(* IEC 61131-3 sources: SortJet_MasterSPS_Aufbau.fbsproj/09_Station/UnterStationsbausteine, 8 files *)

(* ---- Geblaese_Schuetz_FB_V01_00_00.fb.st ---- *)
(* METADATA
{
	"v3Meta": {
		"objectGuid": "c9895c16-daf8-42f8-8f64-ac96a02bd793"
	}
}
*)
FUNCTION_BLOCK Geblaese_Schuetz_FB_V01_00_00
VAR_INPUT

  // BOOLEAN
  bpAktivieren              : BOOL;
  bpStart                   : BOOL;
  bpReset                   : BOOL;
  bpFreigabe                : BOOL;
  bpTeilnehmerErreichbar    : BOOL := TRUE;
  bpIOsBoschDrive               : BOOL;

  // EINGÄNGE
  bpMotorschutzschalter_OK  : BOOL;
  bpDrehzahlErreicht        : BOOL := TRUE; // Sanftanlauf: Drehzahl erreicht (ohne Sanftanlauf TRUE lassen)

  // DROSSELKLAPPE
  bpDrosselklappeAnforderung : BOOL; // Station: Drosselklappe soll offen sein (Transport, Anlegen, Geblaese gestartet)

  // STEUERUNG (wann das Geblaese laufen soll, Aktion Steuerung)
  bpAutomatik        : BOOL;            // Automatik / Check: Geblaese nach Aktivitaet mit Energiesparmodus
  bpAktivitaet       : BOOL;            // Station braucht das Geblaese (z.B. Auftrag aktiv)
  bpAktivitaetFlanke : BOOL;            // Anlegestation: nur die steigende Flanke der Aktivitaet startet, danach Abschaltzeit
  bpTaster           : BOOL;            // Taster am Geblaese: umschalten
  bpHandEin          : BOOL;            // Handbetrieb: Geblaese laeuft, solange gesetzt
  bpSperre           : BOOL;            // Geblaese sofort aus (Reset, Verriegelung)
  tpMindestlaufzeit  : TIME := T#500MS; // Der Taster schaltet erst nach dieser Laufzeit aus

  // STRUKT
  stStationsNummern       : Station_ST;

END_VAR
VAR_OUTPUT

  // BOOLEAN
  bpFehler                 : BOOL;
  bpDone                   : BOOL;
  bpStarteGeblaese         : BOOL; // Geblaese wird angesteuert (Schuetz)
  bpDrosselklappeOeffnen   : BOOL; // Drosselklappe oeffnen: angefordert und Geblaese laeuft

  // WORD
  wpFehlerNr : Fehlerkonstanten_EN;

END_VAR
VAR

  // BOOLEAN
  blErsterZyklus           : BOOL := TRUE; // Initialisierung
  blMeldungAbgesetzt       : BOOL := FALSE;
  blMotorschutzschalter_OK : BOOL;

  // ARRAY
  awlErrorAdditional : ARRAY [0..25]  OF WORD;

  // STEPS
  steplStart      : Steps_TE;

  // TIMER
  tonlStartGeblaese          : TON;
  tonlWarteAufGeblaeseLaeuft : TON;
  toflWarteAufWiederAnlauf   : TOF;
  toflMotorschutz            : TOF;
  toflEnergiesparModus       : TOF; // Energiesparmodus: Geblaese nach der Abschaltzeit ohne Aktivitaet aus
  tonlMindestlaufzeit        : TON;

  // TRIGGER
  rtlAutomatik               : R_TRIG;
  rtlAktivitaet              : R_TRIG;
  rtlTaster                  : R_TRIG;

  // BOOLEAN (Steuerung)
  blTasterAus                : BOOL; // Automatik: Geblaese per Taster ausgeschaltet (bis zur naechsten Aktivitaet)
  blHandTaster               : BOOL; // Handbetrieb: Geblaese per Taster eingeschaltet

END_VAR
VAR

  // HARDWARE EINGAENGE
  in_bMotorschutzschalter_OK    AT %I* : BOOL;

  // HARDWARE AUSGAENGE
  out_bStarteGeblaese           AT %Q* : BOOL;

END_VAR

VAR CONSTANT

  // TIME
  WARTEZEIT_BIS_WIEDERANLAUF          : TIME := T#7000MS;
  WARTEZEIT_BIS_GEBLAESE_HOCHGELAUFEN : TIME := T#2000MS;

END_VAR

//-------------------------------------------------------------------------------------------------
// BAUSTEIN: INITIALISIERUNG
//-------------------------------------------------------------------------------------------------
IF ( blErsterZyklus ) THEN
  blErsterZyklus:=FALSE;

  (* Hinweis:
     - Timer initialisieren
  *)
  toflWarteAufWiederAnlauf(IN:=FALSE);
  tonlWarteAufGeblaeseLaeuft(IN:=FALSE);

END_IF
// IO Zuweisung
IF ( bpIOsBoschDrive ) THEN
  blMotorschutzschalter_OK  := bpMotorschutzschalter_OK;
ELSE
  blMotorschutzschalter_OK  := in_bMotorschutzschalter_OK;
END_IF

//-------------------------------------------------------------------------------------------------
// BAUSTEIN: DEAKTIVIEREN
//-------------------------------------------------------------------------------------------------
IF ( NOT bpAktivieren ) THEN
  bpDone                 := TRUE;
  bpStarteGeblaese       := FALSE;
  bpDrosselklappeOeffnen := FALSE;
  bpFehler   := FALSE;
  wpFehlerNr := cMELDUNG_NULL;

  RETURN;

END_IF

//-------------------------------------------------------------------------------------------------
// BAUSTEIN: STEUERUNG
//-------------------------------------------------------------------------------------------------
Steuerung();

//-------------------------------------------------------------------------------------------------
// BAUSTEIN: TIMER
//-------------------------------------------------------------------------------------------------
toflWarteAufWiederAnlauf(IN :=     out_bStarteGeblaese,
                          PT := WARTEZEIT_BIS_WIEDERANLAUF);

tonlWarteAufGeblaeseLaeuft(IN :=     out_bStarteGeblaese,
                            PT := WARTEZEIT_BIS_GEBLAESE_HOCHGELAUFEN );

toflMotorschutz( IN := blMotorschutzschalter_OK, PT := T#5S );

(* Hinweis:
   - Einschaltverzoegerung
*)
tonlStartGeblaese(IN :=     bpStart
                   AND bpFreigabe
                   AND NOT toflWarteAufWiederAnlauf.Q
                   AND NOT bpReset,
                   PT := T#0S);

//-------------------------------------------------------------------------------------------------
// BAUSTEIN: STEUERUNG
//-------------------------------------------------------------------------------------------------
IF ( bpReset ) THEN

  bpStart   := FALSE;
  bpDone    := FALSE;
  bpReset   := FALSE;
  bpFehler  := FALSE;

  blMeldungAbgesetzt := FALSE;

  wpFehlerNr := cMELDUNG_NULL;

  out_bStarteGeblaese := FALSE;

ELSE
  Start();
  Meldungen();

END_IF

//-------------------------------------------------------------------------------------------------
// BAUSTEIN: AUSGAENGE
//-------------------------------------------------------------------------------------------------
(* Hinweis:
   - Ansteuerung des Geblaeses fuer Stationen, die den Ausgang selbst schalten (z.B. zwei Geblaese oder Ausgang am Umrichter)
   - Die Drosselklappe ist nur offen, wenn sie angefordert ist und das Geblaese laeuft (Drehzahl erreicht)
*)
bpStarteGeblaese       := out_bStarteGeblaese;
bpDrosselklappeOeffnen := bpDrosselklappeAnforderung AND bpDone;
END_FUNCTION_BLOCK

(* ---- Hub_FB_V01_00_00.fb.st ---- *)
(* METADATA
{
	"v3Meta": {
		"objectGuid": "03cf6ff6-d378-4ff5-8445-541e648ef0b8"
	}
}
*)
FUNCTION_BLOCK Hub_FB_V01_00_00
VAR_INPUT

  // BOOLEAN
  bpAktivieren               : BOOL;
  bpStartHubAuf              : BOOL;
  bpStartHubAb               : BOOL;
  bpReset                    : BOOL;
  bpSensorEinlaufNachfolger  : BOOL;
  bpSensorAuslaufVorgaenger  : BOOL;
  bpSensorEinlauf            : BOOL;
  bpSensorAuslauf            : BOOL;

  // STRUCT
  stStationsNummern          : Station_ST;

END_VAR
VAR_OUTPUT

  // BOOLEAN
  bpFehler        : BOOL;
  bpDone          : BOOL;

  // WORD
  wpFehlerNr : Fehlerkonstanten_EN;

  // ENUM
  epHubStatus  : Hub_EN; // Status: Gibt die Aktuelle Position des Antriebs aus

END_VAR

VAR

  // BOOLEAN
  blErsterZyklus        : BOOL := TRUE;

  // TIMER
  tonlMaxWarteZeit                        : TON;
  tonlHubAntriebOK                        : TON;
  tonlMaximaleWartezeitAufReset           : TON;
  tonlFehlermeldungUnterdrueckenAntriebOK : TON;
  tonlReset                               : TON;

  // STEPS
  steplHubAb    : Steps_TE;
  steplHubAuf   : Steps_TE;
  steplReset    : Steps_TE;

END_VAR

VAR
  // HARDWARE EINGÄNGE
  in_bSensorNichtUnten             AT%I* : BOOL;
  in_bSensorNichtOben              AT%I* : BOOL;
  in_bMotorstarter_OK              AT%I* : BOOL;
  in_bLSBremse_OK                  AT%I* : BOOL;
  in_bLS400V_OK                    AT%I* : BOOL;

  // HARDWARE AUSGÄNGE
  out_bHubAbSetzen                 AT%Q* : BOOL;
  out_bHubAufSetzen                AT%Q* : BOOL;
  out_bReset                       AT%Q* : BOOL;
  out_bBremseLoesen                AT%Q* : BOOL;

END_VAR

VAR CONSTANT

  // TIME
  MAXIMALE_WARTEZEIT_HUB                       : TIME := T#5000MS; // Maximale Wartezeit die abgewartet wird bis der Hub-Antrieb auf Position gefahren ist

END_VAR
//-------------------------------------------------------------------------------------------------
// BAUSTEIN: INITIALISIERUNG
//-------------------------------------------------------------------------------------------------
IF ( blErsterZyklus ) THEN
  blErsterZyklus := FALSE;

  (* Hinweis:
     - Timer initialisieren
  *)
  tonlHubAntriebOK(IN:=TRUE);
  tonlMaxWarteZeit(IN:=FALSE);
  tonlFehlermeldungUnterdrueckenAntriebOK( IN := FALSE );

END_IF

//-------------------------------------------------------------------------------------------------
// BAUSTEIN: AKTIONEN
//-------------------------------------------------------------------------------------------------
IF ( bpAktivieren ) THEN

  HubAuf();
  HubAb();

  Ausgaenge();
  Meldungen();
  Timer();
  Reset();

ELSE

  bpDone   := TRUE;
  bpFehler := FALSE;

  IF (bpStartHubAb AND NOT bpStartHubAuf) THEN
    epHubStatus := eHub_Unten;
  ELSIF (bpStartHubAuf AND NOT bpStartHubAb) THEN
    epHubStatus := eHub_Oben;
  ELSIF (bpStartHubAb AND NOT bpStartHubAuf) THEN
    epHubStatus := eHub_Undefiniert;
  END_IF

END_IF
END_FUNCTION_BLOCK

(* ---- Transportsperre_Foerderbaender_FB_V01_00_00.fb.st ---- *)
(* METADATA
{
	"v3Meta": {
		"objectGuid": "85c14a01-ee4c-4a24-bcca-8fef195064c0"
	}
}
*)
{attribute 'excludefrombuild'}
FUNCTION_BLOCK Transportsperre_Foerderbaender_FB_V01_00_00
VAR_INPUT

  // HARDWARE EINGAENGE
  in_bOben            : BOOL; // STATUS: Sensor meldt ausgfahren  [Oben]

  // BOOLEAN
  bpAktivieren        : BOOL;
  bpStartRunter       : BOOL; // BETRIEBTYP: Zylinder wird ausgefahren
  bpStartHoch         : BOOL; // BETRIEBTYP: Zylinder wird eingefahren
  bpReset             : BOOL; // BETRIEBTYP: Zylinderbaustein wird zurueckgesetzt
  bpFreigabe          : BOOL;

  // OPTIONEN
  bpAbfrageObenVorhanden  : BOOL := TRUE;   // Endlagensensor oben vorhanden, sonst gilt die Endlage nach tpBewegungszeit
  bpAbfrageUntenVorhanden : BOOL := TRUE;   // Endlagensensor unten vorhanden, sonst gilt die Endlage nach tpBewegungszeit
  tpBewegungszeit         : TIME := T#800MS; // Bewegungszeit je Richtung ohne Endlagensensor

END_VAR
VAR_OUTPUT

  // BOOLEAN
  bpFehler            : BOOL;
  bpDone              : BOOL;

  // WORD
  wpFehlerNr          : Fehlerkonstanten_EN;

  // ENUM
  wpStatus            : TransportsperrenStatus_EN;

END_VAR
VAR
  // STEPS
  steplHoch         : Steps_TE;
  steplRunter       : Steps_TE;

  // TIMER
  tonlOben                 : TON; // EINSCHALTVERZOEGERUNG: Warten bis der Zylinder eingefahren wurde. Sonst wird ein Fehlerausgegeben
  tonlUnten                : TON; // EINSCHALTVERZOEGERUNG: Warten bis der Zylinder ausgefahren wurde. Sonst wird ein Fehlerausgegeben
  tonlBewegungszeitHoch    : TON; // Bewegungszeit ohne Endlagensensor oben
  tonlBewegungszeitRunter  : TON; // Bewegungszeit ohne Endlagensensor unten
  tofHoch                  : TOF;
  tofRunter                : TOF;

END_VAR

VAR

  // HARDWARE EINGAENGE
  in_bUnten     AT %I* : BOOL; // STATUS: Sensor meldt eingefahren [Unten]

  // HARDWARE AUSGAENGE
  out_bRunter   AT %Q* : BOOL; // AKTION: Zylinder einfahren

END_VAR
VAR CONSTANT

  // TIME
  cZEITLICHE_UEBERWACHUNG_BEWEGUNG_ZYLINDER : TIME := T#15s;

END_VAR
(* Hinweis:
   - Ein Ausgang (Federrueckstell- Ventil): Runter haelt den Ausgang, Hoch nimmt ihn zurueck
*)

//-------------------------------------------------------------------------------------------------
// BAUSTEIN: RESET / DEAKTIVIERT
//-------------------------------------------------------------------------------------------------
(* Hinweis:
   - Reset oder deaktiviert: Ausgang aus, Ketten und Timer zuruecksetzen, Done und Fehler loeschen
   - Der Baustein setzt bpReset selbst zurueck, der Aufrufer wartet nicht auf Done
   - Ein deaktivierter Baustein meldet kein Done; der Aufrufer verknuepft das Warten auf Done
     mit der Aktivierung aus der MK (z.B. Transportsperre.bpDone OR NOT stStationsAufbau.bX)
*)
IF ( bpReset OR NOT bpAktivieren ) THEN

  out_bRunter := FALSE;

  bpStartRunter := FALSE;
  bpStartHoch   := FALSE;

  steplHoch   := STEP_0_E;
  steplRunter := STEP_0_E;

  tonlOben( IN := FALSE );
  tonlUnten( IN := FALSE );
  tonlBewegungszeitHoch( IN := FALSE );
  tonlBewegungszeitRunter( IN := FALSE );
  tofHoch( IN := FALSE );
  tofRunter( IN := FALSE );

  bpDone     := FALSE;
  bpFehler   := FALSE;
  wpFehlerNr := cMELDUNG_NULL;

  bpReset := FALSE;

  RETURN;

END_IF

//-------------------------------------------------------------------------------------------------
// BAUSTEIN: AKTIONEN
//-------------------------------------------------------------------------------------------------
HochFahren();
RunterFahren();

// Umschaltpause zwischen den Richtungen
tofHoch( IN := bpStartHoch, PT := T#1S );
tofRunter( IN := bpStartRunter, PT := T#1S );

//-------------------------------------------------------------------------------------------------
// STATUS DER TRANSPORTSPERRE
//-------------------------------------------------------------------------------------------------
(* Hinweis:
   - Status aus der Sensorik, soweit Endlagensensoren vorhanden sind
   - Ohne Sensor bleibt der Status, den die Schrittketten nach der Bewegungszeit setzen
*)
IF ( bpAbfrageObenVorhanden AND bpAbfrageUntenVorhanden ) THEN

  IF (     in_bOben
       AND NOT in_bUnten )
  THEN
    wpStatus := eTransportsperreOben;
  ELSIF(   in_bUnten
         AND NOT in_bOben )
  THEN
    wpStatus := eTransportsperreUnten;
  ELSE
    wpStatus := eTransportsperreUndefiniert;
  END_IF

ELSIF ( bpAbfrageObenVorhanden ) THEN

  IF ( in_bOben ) THEN
    wpStatus := eTransportsperreOben;
  ELSIF ( wpStatus = eTransportsperreOben ) THEN
    wpStatus := eTransportsperreUndefiniert;
  END_IF

ELSIF ( bpAbfrageUntenVorhanden ) THEN

  IF ( in_bUnten ) THEN
    wpStatus := eTransportsperreUnten;
  ELSIF ( wpStatus = eTransportsperreUnten ) THEN
    wpStatus := eTransportsperreUndefiniert;
  END_IF

END_IF
END_FUNCTION_BLOCK

(* ---- Transportsperre_Kipptisch_FB_V01_00_00.fb.st ---- *)
(* METADATA
{
	"v3Meta": {
		"objectGuid": "32d63b77-62b3-4c1f-9a6d-0b9e7860b01c"
	}
}
*)
{attribute 'excludefrombuild'}
FUNCTION_BLOCK Transportsperre_Kipptisch_FB_V01_00_00
VAR_INPUT

  // BOOLEAN
  bpAktivieren        : BOOL;
  bpStartAusfahren    : BOOL; // BETRIEBTYP: Zylinder wird ausgefahren
  bpStartEinfahren    : BOOL; // BETRIEBTYP: Zylinder wird eingefahren
  bpReset             : BOOL; // BETRIEBTYP: Zylinderbaustein wird zurueckgesetzt
  bpFreigabe          : BOOL; //
  bpFreigabeEinfahren : BOOL; // Freigabe von der Folgestation, dass die Sperre runter fahren darf

  // OPTIONEN
  bpAbfrageAusgefahrenVorhanden : BOOL := TRUE;   // Endlagensensor ausgefahren vorhanden, sonst gilt die Endlage nach tpBewegungszeit
  bpAbfrageEingefahrenVorhanden : BOOL := TRUE;   // Endlagensensor eingefahren vorhanden, sonst gilt die Endlage nach tpBewegungszeit
  tpBewegungszeit               : TIME := T#800MS; // Bewegungszeit je Richtung ohne Endlagensensor

END_VAR
VAR_OUTPUT

  // BOOLEAN
  bpFehler            : BOOL;
  bpDone              : BOOL;
  bpFreigabeKippen    : BOOL;
  bpFreigabeTransport : BOOL;

  // WORD
  wpFehlerNr       : Fehlerkonstanten_EN;

  // ENUM
  wpStatusZylinder : PneumatikZylinderStatus_EN;

END_VAR
VAR
  // STEPS
  steplAusfahren   : Steps_TE;
  steplEinfahren   : Steps_TE;

  // TIMER
  tonlZylinderEingefahren    : TON; // EINSCHALTVERZOEGERUNG: Warten bis der Zylinder eingefahren wurde. Sonst wird ein Fehlerausgegeben
  tonlZylinderAusgefahren    : TON; // EINSCHALTVERZOEGERUNG: Warten bis der Zylinder ausgefahren wurde. Sonst wird ein Fehlerausgegeben
  tonlBewegungszeitEinfahren : TON; // Bewegungszeit ohne Endlagensensor eingefahren
  tonlBewegungszeitAusfahren : TON; // Bewegungszeit ohne Endlagensensor ausgefahren
  tofEinfahren               : TOF;
  tofAusfahren               : TOF;

END_VAR

VAR

  // HARDWARE EINGAENGE
  in_StatusZylinderAusgefahren   AT %I* : BOOL; // STATUS: Sensor meldt ausgfahren  [Oben]
  in_StatusZylinderEingefahren   AT %I* : BOOL; // STATUS: Sensor meldt eingefahren [Unten]

  // HARDWARE AUSGAENGE
  out_ZylinderAusfahren   AT %Q* : BOOL; // AKTION: Zylinder ausfahren
  out_ZylinderEinfahren   AT %Q* : BOOL; // AKTION: Zylinder einfahren

END_VAR
VAR CONSTANT

  // TIME
  cZEITLICHE_UEBERWACHUNG_BEWEGUNG_ZYLINDER : TIME := T#15s;

END_VAR
//-------------------------------------------------------------------------------------------------
// BAUSTEIN: RESET / DEAKTIVIERT
//-------------------------------------------------------------------------------------------------
(* Hinweis:
   - Reset oder deaktiviert: Ausgaenge aus, Ketten und Timer zuruecksetzen, Done und Fehler loeschen
   - Der Baustein setzt bpReset selbst zurueck, der Aufrufer wartet nicht auf Done
   - Ein deaktivierter Zylinder meldet kein Done; der Aufrufer verknuepft das Warten auf Done
     mit der Aktivierung aus der MK (z.B. Zylinder.bpDone OR NOT stStationsAufbau.bX)
*)
IF ( bpReset OR NOT bpAktivieren ) THEN

  out_ZylinderAusfahren := FALSE;
  out_ZylinderEinfahren := FALSE;

  bpStartAusfahren := FALSE;
  bpStartEinfahren := FALSE;

  steplAusfahren := STEP_0_E;
  steplEinfahren := STEP_0_E;

  tonlZylinderAusgefahren( IN := FALSE );
  tonlZylinderEingefahren( IN := FALSE );
  tonlBewegungszeitAusfahren( IN := FALSE );
  tonlBewegungszeitEinfahren( IN := FALSE );
  tofEinfahren( IN := FALSE );
  tofAusfahren( IN := FALSE );

  bpDone              := FALSE;
  bpFehler            := FALSE;
  wpFehlerNr          := cMELDUNG_NULL;
  bpFreigabeKippen    := FALSE;
  bpFreigabeTransport := FALSE;

  bpReset := FALSE;

  RETURN;

END_IF

//-------------------------------------------------------------------------------------------------
// BAUSTEIN: AKTIONEN
//-------------------------------------------------------------------------------------------------
Ausfahren();
Einfahren();

// Umschaltpause zwischen den Richtungen
tofEinfahren( IN := bpStartEinfahren, PT := T#1S );
tofAusfahren( IN := bpStartAusfahren, PT := T#1S );

//-------------------------------------------------------------------------------------------------
// STATUS DES ZYLINDERS
//-------------------------------------------------------------------------------------------------
(* Hinweis:
   - Status aus der Sensorik, soweit Endlagensensoren vorhanden sind
   - Ohne Sensor bleibt der Status, den die Schrittketten nach der Bewegungszeit setzen
*)
IF ( bpAbfrageAusgefahrenVorhanden AND bpAbfrageEingefahrenVorhanden ) THEN

  IF (      in_StatusZylinderAusgefahren
       AND NOT in_StatusZylinderEingefahren )
  THEN
    wpStatusZylinder := eZylinder1Ausgefahren;
  ELSIF(    in_StatusZylinderEingefahren
         AND NOT in_StatusZylinderAusgefahren )
  THEN
    wpStatusZylinder := eZylinder1Eingefahren;
  ELSE
    wpStatusZylinder := eZylinderUndefiniert;
  END_IF

ELSIF ( bpAbfrageAusgefahrenVorhanden ) THEN

  IF ( in_StatusZylinderAusgefahren ) THEN
    wpStatusZylinder := eZylinder1Ausgefahren;
  ELSIF ( wpStatusZylinder = eZylinder1Ausgefahren ) THEN
    wpStatusZylinder := eZylinderUndefiniert;
  END_IF

ELSIF ( bpAbfrageEingefahrenVorhanden ) THEN

  IF ( in_StatusZylinderEingefahren ) THEN
    wpStatusZylinder := eZylinder1Eingefahren;
  ELSIF ( wpStatusZylinder = eZylinder1Eingefahren ) THEN
    wpStatusZylinder := eZylinderUndefiniert;
  END_IF

END_IF

bpFreigabeKippen    := ( wpStatusZylinder = eZylinder1Ausgefahren );
bpFreigabeTransport := ( wpStatusZylinder = eZylinder1Eingefahren );
END_FUNCTION_BLOCK

(* ---- Wandverstellung_FB_V01_00_00.fb.st ---- *)
(* METADATA
{
	"v3Meta": {
		"objectGuid": "10dab8d5-0a44-4f93-9a62-9b59bb1a4144"
	}
}
*)
{attribute 'excludefrombuild'}
FUNCTION_BLOCK Wandverstellung_FB_V01_00_00
VAR_INPUT

  // BOOLEAN
  bpWandverstellungOeffnen    : BOOL;
  bpWandverstellungSchliessen : BOOL;
  bpReset                     : BOOL;
  bpAktivieren                : BOOL;

  // OPTIONEN
  bpAbfrageGeoeffnetVorhanden   : BOOL := TRUE;   // Endlagensensoren geoeffnet vorhanden, sonst gilt die Endlage nach tpBewegungszeit
  bpAbfrageGeschlossenVorhanden : BOOL := TRUE;   // Endlagensensoren geschlossen vorhanden, sonst gilt die Endlage nach tpBewegungszeit
  tpBewegungszeit               : TIME := T#800MS; // Bewegungszeit je Richtung ohne Endlagensensor

END_VAR
VAR_OUTPUT

  // BOOLEAN
  bpDone    : BOOL;
  bpFehler  : BOOL;

  // WORD
  wpFehlerNr  : Fehlerkonstanten_EN;

  // ENUM
  epWandStatus  : WandOeffnung_EN;// Status: Gibt die Aktuelle Position des Antriebs aus

END_VAR
VAR

  // STEPS
  steplWandverstellungOeffnen    : Steps_TE;
  steplWandverstellungSchliessen : Steps_TE;

  // TIMER
  tonlEingefahrenWandEinlaufseite  : TON; // EINSCHALTVERZOEGERUNG: Warten bis der Zylinder verfahren wurde. Sonst wird ein Fehlerausgegeben
  tonlAusgefahrenWandEinlaufseite  : TON; // EINSCHALTVERZOEGERUNG: Warten bis der Zylinder verfahren wurde. Sonst wird ein Fehlerausgegeben
  tonlEingefahrenWandAuslaufseite  : TON; // EINSCHALTVERZOEGERUNG: Warten bis der Zylinder verfahren wurde. Sonst wird ein Fehlerausgegeben
  tonlAusgefahrenWandAuslaufseite  : TON; // EINSCHALTVERZOEGERUNG: Warten bis der Zylinder verfahren wurde. Sonst wird ein Fehlerausgegeben
  tonlBewegungszeitOeffnen         : TON; // Bewegungszeit ohne Endlagensensor geoeffnet
  tonlBewegungszeitSchliessen      : TON; // Bewegungszeit ohne Endlagensensor geschlossen

END_VAR
VAR

  // HARDWARE EINGAENGE
  in_bWandEinlaufseiteGeoeffnet    AT %I* : BOOL; // STATUS: Sensor meldet geöffnet
  in_bWandEinlaufseiteGeschlossen  AT %I* : BOOL; // STATUS: Sensor meldet geschlossen
  in_bWandAuslaufseiteGeoeffnet    AT %I* : BOOL; // STATUS: Sensor meldet geöffnet
  in_bWandAuslaufseiteGeschlossen  AT %I* : BOOL; // STATUS: Sensor meldet geschlossen

  // HARDWARE AUSGAENGE
  out_bWandverstellungOeffnen      AT %Q* : BOOL; // AKTION: Verstellen der Wandoeffnung -> Maximal Geoeffnet
  out_bWandverstellungSchliessen   AT %Q* : BOOL; // AKTION: Verstellen der Wandoeffnung -> Minimal Geoeffnet

END_VAR

//-------------------------------------------------------------------------------------------------
// BAUSTEIN: RESET / DEAKTIVIERT
//-------------------------------------------------------------------------------------------------
(* Hinweis:
   - Reset oder deaktiviert: Ausgaenge aus, Ketten und Timer zuruecksetzen, Done und Fehler loeschen
   - Der Baustein setzt bpReset selbst zurueck, der Aufrufer wartet nicht auf Done
   - Ein deaktivierter Baustein meldet kein Done; der Aufrufer verknuepft das Warten auf Done
     mit der Aktivierung aus der MK (z.B. Wandverstellung.bpDone OR NOT stStationsAufbau.bX)
*)
IF ( bpReset OR NOT bpAktivieren ) THEN

  out_bWandverstellungOeffnen    := FALSE;
  out_bWandverstellungSchliessen := FALSE;

  bpWandverstellungOeffnen    := FALSE;
  bpWandverstellungSchliessen := FALSE;

  steplWandverstellungOeffnen    := STEP_0_E;
  steplWandverstellungSchliessen := STEP_0_E;

  tonlEingefahrenWandEinlaufseite( IN := FALSE );
  tonlAusgefahrenWandEinlaufseite( IN := FALSE );
  tonlEingefahrenWandAuslaufseite( IN := FALSE );
  tonlAusgefahrenWandAuslaufseite( IN := FALSE );
  tonlBewegungszeitOeffnen( IN := FALSE );
  tonlBewegungszeitSchliessen( IN := FALSE );

  wpFehlerNr := cMELDUNG_NULL;
  bpFehler   := FALSE;
  bpDone     := FALSE;

  bpReset := FALSE;

  RETURN;

END_IF

//-------------------------------------------------------------------------------------------------
// BAUSTEIN: AKTIONEN
//-------------------------------------------------------------------------------------------------
WandverstellungOeffnen();
WandverstellungSchliessen();

//-------------------------------------------------------------------------------------------------
// STATUS DER WAND
//-------------------------------------------------------------------------------------------------
(* Hinweis:
   - Status aus der Sensorik, soweit Endlagensensoren vorhanden sind (beide Seiten)
   - Ohne Sensor bleibt der Status, den die Schrittketten nach der Bewegungszeit setzen
*)
IF ( bpAbfrageGeoeffnetVorhanden AND bpAbfrageGeschlossenVorhanden ) THEN

  IF (     in_bWandEinlaufseiteGeschlossen AND in_bWandAuslaufseiteGeschlossen
       AND NOT in_bWandEinlaufseiteGeoeffnet AND NOT in_bWandAuslaufseiteGeoeffnet )
  THEN
    epWandStatus := eWandOeffnung_Geschlossen;
  ELSIF (     in_bWandEinlaufseiteGeoeffnet AND in_bWandAuslaufseiteGeoeffnet
          AND NOT in_bWandEinlaufseiteGeschlossen AND NOT in_bWandAuslaufseiteGeschlossen )
  THEN
    epWandStatus := eWandOeffnung_Offen;
  ELSE
    epWandStatus := eWandOeffnung_Undefiniert;
  END_IF

ELSIF ( bpAbfrageGeoeffnetVorhanden ) THEN

  IF ( in_bWandEinlaufseiteGeoeffnet AND in_bWandAuslaufseiteGeoeffnet ) THEN
    epWandStatus := eWandOeffnung_Offen;
  ELSIF ( epWandStatus = eWandOeffnung_Offen ) THEN
    epWandStatus := eWandOeffnung_Undefiniert;
  END_IF

ELSIF ( bpAbfrageGeschlossenVorhanden ) THEN

  IF ( in_bWandEinlaufseiteGeschlossen AND in_bWandAuslaufseiteGeschlossen ) THEN
    epWandStatus := eWandOeffnung_Geschlossen;
  ELSIF ( epWandStatus = eWandOeffnung_Geschlossen ) THEN
    epWandStatus := eWandOeffnung_Undefiniert;
  END_IF

END_IF
END_FUNCTION_BLOCK

(* ---- ZylinderPneumatik_3Wege_FB_V01_00_00.fb.st ---- *)
(* METADATA
{
	"v3Meta": {
		"objectGuid": "530c17d7-3762-455b-8431-d2a354444d9d"
	}
}
*)
FUNCTION_BLOCK ZylinderPneumatik_3Wege_FB_V01_00_00
VAR_INPUT

  // BOOLEAN
  blErsterZyklus              : BOOL;
  bpAktivieren                : BOOL;
  bpFreigabe                  : BOOL; // FREIGABE Pneumatik: ohne Freigabe Ventile aus, Bewegung pausiert (Startbefehl bleibt erhalten)
  bpStartPneumatik            : BOOL; // Starten der Zylinder
  bpReset                     : BOOL; // BETRIEBTYP: Zylinderbaustein wird zurueckgesetzt
  bpZylinderAbfragenVorhanden : BOOL := TRUE;  // Hinweis: Manche Zylinder haben keine Abfragen
  bpEinAusFahrenLogikDrehen   : BOOL := FALSE; // Hinweis: Manche Zylinder haben keine Abfragen
  tpWartezeitOhneAbfrage      : TIME := T#1S;  // Hinweis: Ohne Abfragen gilt die Stellung nach dieser Zeit als erreicht
  bpZweiterZylinderVorhanden  : BOOL := TRUE;  // Hinweis: Mit nur einem Zylinder (z.B. Rollenleiste) sind die Signale von Zylinder 2 ohne Funktion, es gibt nur Geschlossen (16 mm) und Geoeffnet (29 mm)

  // ENUM
  epOeffnungsStellung  : PneumatikZylinderStatus_EN;

END_VAR

VAR_OUTPUT

  // BOOLEAN
  bpFehler                       : BOOL;
  bpDone                         : BOOL;

  // WORD
  wpFehlerNr                     : Fehlerkonstanten_EN;

  // ENUM
  wpStatusZylinder               : PneumatikZylinderStatus_EN;

END_VAR
VAR

  // HARDWARE EINGAENGE
  in_bStatusZylinder1Ausgefahren   AT %I* : BOOL; // STATUS: Sensor meldet ausgfahren
  in_bStatusZylinder1Eingefahren   AT %I* : BOOL; // STATUS: Sensor meldet eingefahren
  in_bStatusZylinder2Ausgefahren   AT %I* : BOOL; // STATUS: Sensor meldet ausgfahren
  in_bStatusZylinder2Eingefahren   AT %I* : BOOL; // STATUS: Sensor meldet eingefahren

  // HARDWARE AUSGAENGE
  out_bZylinder1Ausfahren   AT %Q* : BOOL; // AKTION: Zylinder 1 ausfahren
  out_bZylinder1Einfahren   AT %Q* : BOOL; // AKTION: Zylinder 1 einfahren
  out_bZylinder2Ausfahren   AT %Q* : BOOL; // AKTION: Zylinder 2 ausfahren
  out_bZylinder2Einfahren   AT %Q* : BOOL; // AKTION: Zylinder 2 einfahren

  // BOOLEAN
  blZylinder2Ausgefahren : BOOL; // Zylinder 2 ausgefahren, bei nur einem Zylinder folgt das Signal Zylinder 1
  blZylinder2Eingefahren : BOOL; // Zylinder 2 eingefahren, bei nur einem Zylinder folgt das Signal Zylinder 1

  // ENUM
  elStellung : PneumatikZylinderStatus_EN; // Wirksame Sollstellung (Geschlossen = 16 mm, Geoeffnet = 29 mm, ein Zylinder: 23 mm = 29 mm)

  // STEPS
  steplAusfahren   : Steps_TE;

  // TIMER
  tonlZylinder1Eingefahren  : TON; // EINSCHALTVERZOEGERUNG: Warten bis der Zylinder eingefahren wurde. Sonst wird ein Fehlerausgegeben
  tonlZylinder1Ausgefahren  : TON; // EINSCHALTVERZOEGERUNG: Warten bis der Zylinder ausgefahren wurde. Sonst wird ein Fehlerausgegeben
  tonlZylinder2Eingefahren  : TON; // EINSCHALTVERZOEGERUNG: Warten bis der Zylinder eingefahren wurde. Sonst wird ein Fehlerausgegeben
  tonlZylinder2Ausgefahren  : TON; // EINSCHALTVERZOEGERUNG: Warten bis der Zylinder ausgefahren wurde. Sonst wird ein Fehlerausgegeben
  tonlWarteZeitAufVentile   : TON; // EINSCHALTVERZOEGERUNG: wenn keine Abfragen verbaut sind, pauschal die Schaltung der Ventile zurücksetzen

END_VAR
//-------------------------------------------------------------------------------------------------
// INITIALISIERUNG
//-------------------------------------------------------------------------------------------------
IF ( blErsterZyklus  ) THEN
  blErsterZyklus := FALSE;
  epOeffnungsStellung := eZylinderStellung16mm;
END_IF

//-------------------------------------------------------------------------------------------------
// BAUSTEIN: RESET / DEAKTIVIERT
//-------------------------------------------------------------------------------------------------
(* Hinweis:
   - Reset oder deaktiviert: Ausgaenge aus, Kette und Timer zuruecksetzen, Done und Fehler loeschen
   - Der Baustein setzt bpReset selbst zurueck, der Aufrufer wartet nicht auf Done
   - Ein deaktivierter Zylinder meldet kein Done; der Aufrufer verknuepft das Warten auf Done
     mit der Aktivierung aus der MK (z.B. Zylinder.bpDone OR NOT stStationsAufbau.bX)
*)
IF ( bpReset OR NOT bpAktivieren ) THEN

  out_bZylinder1Ausfahren := FALSE;
  out_bZylinder1Einfahren := FALSE;
  out_bZylinder2Ausfahren := FALSE;
  out_bZylinder2Einfahren := FALSE;

  bpStartPneumatik := FALSE;

  steplAusfahren := STEP_0_E;

  tonlZylinder1Ausgefahren( IN := FALSE );
  tonlZylinder1Eingefahren( IN := FALSE );
  tonlZylinder2Ausgefahren( IN := FALSE );
  tonlZylinder2Eingefahren( IN := FALSE );
  tonlWarteZeitAufVentile( IN := FALSE );

  bpDone     := FALSE;
  bpFehler   := FALSE;
  wpFehlerNr := cMELDUNG_NULL;

  bpReset := FALSE;

  RETURN;

END_IF

//-------------------------------------------------------------------------------------------------
// AKTIONEN
//-------------------------------------------------------------------------------------------------
(* Hinweis:
   - Mit nur einem Zylinder folgen die Signale von Zylinder 2 denen von Zylinder 1
*)
IF ( bpZweiterZylinderVorhanden ) THEN
  blZylinder2Ausgefahren := in_bStatusZylinder2Ausgefahren;
  blZylinder2Eingefahren := in_bStatusZylinder2Eingefahren;
ELSE
  blZylinder2Ausgefahren := in_bStatusZylinder1Ausgefahren;
  blZylinder2Eingefahren := in_bStatusZylinder1Eingefahren;
END_IF

(* Hinweis Freigabe Pneumatik:
   - Ohne Freigabe: Ventile aus, Kette und Ueberwachungszeiten zuruecksetzen (kein Timeout-Fehler)
   - Der Startbefehl bleibt erhalten: kommt die Freigabe zurueck, wird die Bewegung neu gestartet
*)
IF NOT bpFreigabe THEN
  out_bZylinder1Ausfahren := FALSE;
  out_bZylinder1Einfahren := FALSE;
  out_bZylinder2Ausfahren := FALSE;
  out_bZylinder2Einfahren := FALSE;
  steplAusfahren := STEP_0_E;
  tonlZylinder1Ausgefahren( IN := FALSE );
  tonlZylinder1Eingefahren( IN := FALSE );
  tonlZylinder2Ausgefahren( IN := FALSE );
  tonlZylinder2Eingefahren( IN := FALSE );
  tonlWarteZeitAufVentile( IN := FALSE );
  bpDone := FALSE;
ELSE
  AusEinFahren();
END_IF

//-------------------------------------------------------------------------------------------------
// STATUS DER ZYLINDER
//-------------------------------------------------------------------------------------------------
(* Hinweis:
   - Status aus der Sensorik, wenn Abfragen vorhanden sind
   - Ohne Abfragen bleibt der Status, den die Schrittkette nach der Wartezeit setzt
*)
IF ( bpZylinderAbfragenVorhanden ) THEN

  IF NOT bpEinAusFahrenLogikDrehen THEN

    IF ( in_bStatusZylinder1Ausgefahren ) THEN
      IF (blZylinder2Ausgefahren) THEN
        wpStatusZylinder := eZylinderStellung29mm;
      ELSE
        wpStatusZylinder := eZylinderStellung23mm;
      END_IF

    ELSE
      IF (blZylinder2Ausgefahren) THEN
        wpStatusZylinder := eZylinderStellung23mm;
      ELSE
        wpStatusZylinder := eZylinderStellung16mm;
      END_IF
    END_IF

  ELSE

    IF in_bStatusZylinder1Eingefahren THEN

      IF (blZylinder2Eingefahren) THEN
        wpStatusZylinder := eZylinderStellung29mm;
      ELSE
        wpStatusZylinder := eZylinderStellung23mm;
      END_IF

    ELSE

      IF (blZylinder2Eingefahren) THEN
        wpStatusZylinder := eZylinderStellung23mm;
      ELSE
        wpStatusZylinder := eZylinderStellung16mm;
      END_IF

    END_IF

  END_IF

END_IF
END_FUNCTION_BLOCK

(* ---- ZylinderPneumatik_FB_V01_00_00.fb.st ---- *)
(* METADATA
{
	"v3Meta": {
		"objectGuid": "c49e37bf-a253-4691-9610-12ec51ad1d15"
	}
}
*)
FUNCTION_BLOCK ZylinderPneumatik_FB_V01_00_00
VAR_INPUT

  // BOOLEAN
  bpReset            : BOOL;
  bpAktivieren       : BOOL;

  bpFreigabe         : BOOL; // FREIGABE Pneumatik: ohne Freigabe Ventile aus, Bewegung pausiert (Startbefehl bleibt erhalten)
  bpStartAusfahren   : BOOL; // BETRIEBTYP: Zylinder wird ausgefahren
  bpStartEinfahren   : BOOL; // BETRIEBTYP: Zylinder wird eingefahren

  // OPTIONEN
  bpAbfrageAusgefahrenVorhanden : BOOL := TRUE;   // Endlagensensor ausgefahren vorhanden, sonst gilt die Endlage nach tpBewegungszeit
  bpAbfrageEingefahrenVorhanden : BOOL := TRUE;   // Endlagensensor eingefahren vorhanden, sonst gilt die Endlage nach tpBewegungszeit
  bpAbfrageAusgefahrenOeffner   : BOOL := FALSE;   // Endlagensensor ausgefahren vorhanden, sonst gilt die Endlage nach tpBewegungszeit
  bpAbfrageEingefahrenOeffner   : BOOL := FALSE;   // Endlagensensor eingefahren vorhanden, sonst gilt die Endlage nach tpBewegungszeit
  tpBewegungszeit               : TIME := T#1S; // Bewegungszeit je Richtung ohne Endlagensensor

  // HARDWARE EINGAENGE
  in_bStatusZylinderAusgefahren   : BOOL; // STATUS: Sensor meldt ausgefahren  [Oben]
  in_bStatusZylinderEingefahren   : BOOL; // STATUS: Sensor meldt eingefahren [Unten]

END_VAR
VAR_OUTPUT

  // BOOLEAN
  bpFehler                       : BOOL;
  bpDone                         : BOOL;

  // WORD
  wpFehlerNr       : Fehlerkonstanten_EN;

  // ENUM
  epStatusZylinder : PneumatikZylinderStatus_EN;

END_VAR
VAR

  // STEPS
  steplAusfahren   : Steps_TE;
  steplEinfahren   : Steps_TE;

  // TIMER
  tonZylinderEingefahren     : TON; // EINSCHALTVERZOEGERUNG: Warten bis der Zylinder eingefahren wurde. Sonst wird ein Fehlerausgegeben
  tonZylinderAusgefahren     : TON; // EINSCHALTVERZOEGERUNG: Warten bis der Zylinder ausgefahren wurde. Sonst wird ein Fehlerausgegeben
  tonlBewegungszeitEinfahren : TON; // Bewegungszeit ohne Endlagensensor eingefahren
  tonlBewegungszeitAusfahren : TON; // Bewegungszeit ohne Endlagensensor ausgefahren

END_VAR
VAR

  // HARDWARE AUSGAENGE
  out_bZylinderAusfahren    : BOOL; // AKTION: Zylinder ausfahren
  out_bZylinderEinfahren    : BOOL; // AKTION: Zylinder einfahren

END_VAR
VAR CONSTANT

  // TIME
  cZEITLICHE_UEBERWACHUNG_BEWEGUNG_ZYLINDER : TIME := T#15s;

END_VAR
//-------------------------------------------------------------------------------------------------
// BAUSTEIN: RESET / DEAKTIVIERT
//-------------------------------------------------------------------------------------------------
(* Hinweis:
   - Reset oder deaktiviert: Ausgaenge aus, Ketten und Timer zuruecksetzen, Done und Fehler loeschen
   - Ein deaktivierter Zylinder meldet kein Done; der Aufrufer verknuepft das Warten auf Done
     mit der Aktivierung aus der MK (z.B. Zylinder.bpDone OR NOT stStationsAufbau.bX)
*)
IF ( bpReset OR NOT bpAktivieren ) THEN

  out_bZylinderAusfahren := FALSE;
  out_bZylinderEinfahren := FALSE;

  bpStartAusfahren := FALSE;
  bpStartEinfahren := FALSE;

  steplAusfahren := STEP_0_E;
  steplEinfahren := STEP_0_E;

  tonZylinderAusgefahren( IN := FALSE );
  tonZylinderEingefahren( IN := FALSE );
  tonlBewegungszeitAusfahren( IN := FALSE );
  tonlBewegungszeitEinfahren( IN := FALSE );

  bpDone           := FALSE;
  bpFehler         := FALSE;
  wpFehlerNr       := cMELDUNG_NULL;

  bpReset := FALSE;

  RETURN;

END_IF

IF bpAbfrageEingefahrenOeffner THEN
  in_bStatusZylinderEingefahren := NOT in_bStatusZylinderEingefahren;
END_IF
IF bpAbfrageAusgefahrenOeffner THEN
  in_bStatusZylinderAusgefahren := NOT in_bStatusZylinderAusgefahren;
END_IF

//-------------------------------------------------------------------------------------------------
// BAUSTEIN: AKTIONEN
//-------------------------------------------------------------------------------------------------
(* Hinweis Freigabe Pneumatik:
   - Ohne Freigabe: Ventile aus, Ketten und Ueberwachungszeiten zuruecksetzen (kein Timeout-Fehler)
   - Der Startbefehl bleibt erhalten: kommt die Freigabe zurueck, wird die Bewegung neu gestartet
*)
IF NOT bpFreigabe THEN
  out_bZylinderAusfahren := FALSE;
  out_bZylinderEinfahren := FALSE;
  steplAusfahren := STEP_0_E;
  steplEinfahren := STEP_0_E;
  tonZylinderAusgefahren( IN := FALSE );
  tonZylinderEingefahren( IN := FALSE );
  tonlBewegungszeitAusfahren( IN := FALSE );
  tonlBewegungszeitEinfahren( IN := FALSE );
  bpDone := FALSE;
ELSE
  Ausfahren();
  Einfahren();
END_IF

//-------------------------------------------------------------------------------------------------
// STATUS DES ZYLINDERS
//-------------------------------------------------------------------------------------------------
(* Hinweis:
   - Status aus der Sensorik, soweit Endlagensensoren vorhanden sind
   - Ohne Sensor bleibt der Status, den die Schrittketten nach der Bewegungszeit setzen
*)
IF ( bpAbfrageAusgefahrenVorhanden AND bpAbfrageEingefahrenVorhanden ) THEN

  IF (      in_bStatusZylinderAusgefahren
       AND NOT in_bStatusZylinderEingefahren )
  THEN
    epStatusZylinder := eZylinderAusgefahren;
  ELSIF(    in_bStatusZylinderEingefahren
         AND NOT in_bStatusZylinderAusgefahren )
  THEN
    epStatusZylinder := eZylinderEingefahren;
  ELSE
    epStatusZylinder := eZylinderUndefiniert;
  END_IF

ELSIF ( bpAbfrageAusgefahrenVorhanden ) THEN

  IF ( in_bStatusZylinderAusgefahren ) THEN
    epStatusZylinder := eZylinderAusgefahren;
  ELSIF ( epStatusZylinder = eZylinderAusgefahren ) THEN
    epStatusZylinder := eZylinderUndefiniert;
  END_IF

ELSIF ( bpAbfrageEingefahrenVorhanden ) THEN

  IF ( in_bStatusZylinderEingefahren ) THEN
    epStatusZylinder := eZylinderEingefahren;
  ELSIF ( epStatusZylinder = eZylinderEingefahren ) THEN
    epStatusZylinder := eZylinderUndefiniert;
  END_IF

END_IF
END_FUNCTION_BLOCK

(* ---- ZylinderPneumatik_Federrueck_FB_V01_00_00.fb.st ---- *)
(* METADATA
{
	"v3Meta": {
		"objectGuid": "b2af587c-0d32-447c-a5c9-96380651afc9"
	}
}
*)
FUNCTION_BLOCK ZylinderPneumatik_Federrueck_FB_V01_00_00
VAR_INPUT

  // BOOLEAN
  bpAktivieren     : BOOL;
  bpFreigabe       : BOOL; // FREIGABE Pneumatik: ohne Freigabe Ventil aus (Feder faehrt zurueck), Bewegung pausiert (Startbefehl bleibt erhalten)
  bpStartAusfahren : BOOL; // BETRIEBTYP: Zylinder wird ausgefahren
  bpStartEinfahren : BOOL; // BETRIEBTYP: Zylinder wird eingefahren
  bpReset          : BOOL; // BETRIEBTYP: Zylinderbaustein wird zurueckgesetzt

  // OPTIONEN
  bpAbfrageAusgefahrenVorhanden : BOOL := TRUE;   // Endlagensensor ausgefahren vorhanden, sonst gilt die Endlage nach tpBewegungszeit
  bpAbfrageEingefahrenVorhanden : BOOL := TRUE;   // Endlagensensor eingefahren vorhanden, sonst gilt die Endlage nach tpBewegungszeit
  tpBewegungszeit               : TIME := T#800MS; // Bewegungszeit je Richtung ohne Endlagensensor

END_VAR
VAR_OUTPUT

  // BOOLEAN
  bpFehler   : BOOL;
  bpDone     : BOOL;

  // WORD
  wpFehlerNr : Fehlerkonstanten_EN;

  // ENUM
  epStatusZylinder : PneumatikZylinderStatus_EN;

END_VAR
VAR

  // HARDWARE EINGAENGE
  in_bStatusZylinderAusgefahren   AT %I* : BOOL; // STATUS: Sensor meldt ausgfahren
  in_bStatusZylinderEingefahren   AT %I* : BOOL; // STATUS: Sensor meldt eingefahren

  // HARDWARE AUSGAENGE
  out_bZylinderAusfahren          AT %Q* : BOOL; // AUSGANG: (in Glasflussrichtung) Signal zum Ausfahren  [Federrueckstell- Ventiel]

  // STEPS
  steplAusfahren   : Steps_TE;
  steplEinfahren   : Steps_TE;

  // TIMER
  tonlZylinderEingefahren    : TON; // EINSCHALTVERZOEGERUNG: Warten bis der Zylinder eingefahren wurde. Sonst wird ein Fehlerausgegeben
  tonlZylinderAusgefahren    : TON; // EINSCHALTVERZOEGERUNG: Warten bis der Zylinder ausgefahren wurde. Sonst wird ein Fehlerausgegeben
  tonlBewegungszeitEinfahren : TON; // Bewegungszeit ohne Endlagensensor eingefahren
  tonlBewegungszeitAusfahren : TON; // Bewegungszeit ohne Endlagensensor ausgefahren

END_VAR
VAR CONSTANT

  // TIME
  cZEITLICHE_UEBERWACHUNG_BEWEGUNG_ZYLINDER : TIME := T#5s;

END_VAR
(* Hinweis:
   - Es handelt sich bei diesem Baustein um eine Ansteuerung fuer ein Federrueckstell- Ventiel
     => Der Ausgang bleibt nach dem Ausfahren gesetzt, Einfahren nimmt ihn zurueck
*)

//-------------------------------------------------------------------------------------------------
// BAUSTEIN: RESET / DEAKTIVIERT
//-------------------------------------------------------------------------------------------------
(* Hinweis:
   - Reset oder deaktiviert: Ausgang aus, Ketten und Timer zuruecksetzen, Done und Fehler loeschen
   - Der Baustein setzt bpReset selbst zurueck, der Aufrufer wartet nicht auf Done
   - Ein deaktivierter Zylinder meldet kein Done; der Aufrufer verknuepft das Warten auf Done
     mit der Aktivierung aus der MK (z.B. Zylinder.bpDone OR NOT stStationsAufbau.bX)
*)
IF ( bpReset OR NOT bpAktivieren ) THEN

  out_bZylinderAusfahren := FALSE;

  bpStartAusfahren := FALSE;
  bpStartEinfahren := FALSE;

  steplAusfahren := STEP_0_E;
  steplEinfahren := STEP_0_E;

  tonlZylinderAusgefahren( IN := FALSE );
  tonlZylinderEingefahren( IN := FALSE );
  tonlBewegungszeitAusfahren( IN := FALSE );
  tonlBewegungszeitEinfahren( IN := FALSE );

  bpDone     := FALSE;
  bpFehler   := FALSE;
  wpFehlerNr := cMELDUNG_NULL;

  bpReset := FALSE;

  RETURN;

END_IF

//-------------------------------------------------------------------------------------------------
// BAUSTEIN: AKTIONEN
//-------------------------------------------------------------------------------------------------
(* Hinweis Freigabe Pneumatik:
   - Ohne Freigabe: Ventil aus, Ketten und Ueberwachungszeiten zuruecksetzen (kein Timeout-Fehler)
   - Der Startbefehl bleibt erhalten: kommt die Freigabe zurueck, wird die Bewegung neu gestartet
*)
IF NOT bpFreigabe THEN
  out_bZylinderAusfahren := FALSE;
  steplAusfahren := STEP_0_E;
  steplEinfahren := STEP_0_E;
  tonlZylinderAusgefahren( IN := FALSE );
  tonlZylinderEingefahren( IN := FALSE );
  tonlBewegungszeitAusfahren( IN := FALSE );
  tonlBewegungszeitEinfahren( IN := FALSE );
  bpDone := FALSE;
ELSE
  Ausfahren();
  Einfahren();
END_IF

//-------------------------------------------------------------------------------------------------
// STATUS DES ZYLINDERS
//-------------------------------------------------------------------------------------------------
(* Hinweis:
   - Status aus der Sensorik, soweit Endlagensensoren vorhanden sind
   - Ohne Sensor bleibt der Status, den die Schrittketten nach der Bewegungszeit setzen
*)
IF ( bpAbfrageAusgefahrenVorhanden AND bpAbfrageEingefahrenVorhanden ) THEN

  IF (      in_bStatusZylinderAusgefahren
       AND NOT in_bStatusZylinderEingefahren )
  THEN
    epStatusZylinder := eZylinderAusgefahren;
  ELSIF(    in_bStatusZylinderEingefahren
         AND NOT in_bStatusZylinderAusgefahren )
  THEN
    epStatusZylinder := eZylinderEingefahren;
  ELSE
    epStatusZylinder := eZylinderUndefiniert;
  END_IF

ELSIF ( bpAbfrageAusgefahrenVorhanden ) THEN

  IF ( in_bStatusZylinderAusgefahren ) THEN
    epStatusZylinder := eZylinderAusgefahren;
  ELSIF ( epStatusZylinder = eZylinderAusgefahren ) THEN
    epStatusZylinder := eZylinderUndefiniert;
  END_IF

ELSIF ( bpAbfrageEingefahrenVorhanden ) THEN

  IF ( in_bStatusZylinderEingefahren ) THEN
    epStatusZylinder := eZylinderEingefahren;
  ELSIF ( epStatusZylinder = eZylinderEingefahren ) THEN
    epStatusZylinder := eZylinderUndefiniert;
  END_IF

END_IF
END_FUNCTION_BLOCK
